TYPE ST_Error :
STRUCT
	nSource:		UDINT;
	nType:			UDINT;
	sMsg:			STRING(80);
END_STRUCT
END_TYPE

(* stored: Version 1.1.0.1, ProductVersion 3.1.4024.12
   DUT ST_Error: Id {48592411-e712-4fc5-bcf1-87b513435750} *)
